(* IEC 61131-3 sources: twincat-st/tests/fixtures/negative, 10 files *)

(* ---- cp8_change_detect.st ---- *)
FUNCTION_BLOCK FB_ChangeDetect
VAR_INPUT
  fSetpoint  : LREAL;  // [mm]
  bStart    : BOOL;
END_VAR
VAR_OUTPUT
  bSetpointChanged : BOOL;
END_VAR
VAR
  fTarget    : LREAL;  // [mm] setpoint latched at start
END_VAR
IF bStart THEN
  fTarget := fSetpoint;
END_IF
bSetpointChanged := (fTarget <> fSetpoint);
END_FUNCTION_BLOCK

(* ---- FB_AbstractHook.st ---- *)
// CP24 must stay quiet on the abstract method's parameter: it has no body to use
// it in, by design. The concrete method's parameter is used and also stays quiet.
FUNCTION_BLOCK ABSTRACT FB_AbstractHook
VAR_OUTPUT
    nLast : INT;
END_VAR

METHOD ABSTRACT OnStep
VAR_INPUT
    nStep : INT;
END_VAR

METHOD Record
VAR_INPUT
    nValue : INT;
END_VAR
nLast := nValue;

(* ---- FB_ConditionalCallsClean.st ---- *)
// X12, CP7 and CP12 must stay quiet on every shape here. A timer reset with
// IN := FALSE on the way into its state, blocks called unconditionally, an Error
// bound with '=>', read as a member, or handed on whole, and an output written in
// both branches of one IF are all correct.
FUNCTION_BLOCK FB_ConditionalCallsClean
VAR_INPUT
    bStart   : BOOL;
    bSensor  : BOOL;
    fPos     : LREAL;    // mm
END_VAR
VAR_OUTPUT
    bFault   : BOOL;
END_VAR
VAR
    eStep    : E_Step;
    tonWait  : TON;
    tonStep  : TON;
    fbEdge   : R_TRIG;
    fbMove   : MC_MoveAbsolute;
    fbPower  : MC_Power;
    fbHome   : MC_Home;
    axisX    : AXIS_REF;
    bMoveErr : BOOL;
    qbValve AT %Q* : BOOL;
END_VAR
fbEdge(CLK := bSensor);
tonStep(IN := eStep = E_Step.Settle, PT := T#500MS);
CASE eStep OF
    E_Step.Idle:
        IF bStart THEN
            tonWait(IN := FALSE);   // lint:allow CP20 the reset on the way into Wait
            eStep := E_Step.Wait;
        END_IF
    E_Step.Wait:
        tonWait(IN := TRUE, PT := T#2S);
        IF tonWait.Q OR fbEdge.Q THEN
            eStep := E_Step.Settle;
        END_IF
    E_Step.Settle:
        IF tonStep.Q THEN
            eStep := E_Step.Idle;
        END_IF
    E_Step.Error:
        eStep := E_Step.Idle;
ELSE
    eStep := E_Step.Error;
END_CASE
fbPower(Axis := axisX, Enable := TRUE);
fbMove(Axis := axisX, Execute := eStep = E_Step.Settle, Position := fPos,
       Velocity := 50.0, Error => bMoveErr);
fbHome(Axis := axisX, Execute := bStart);
IF bMoveErr OR fbPower.Error THEN
    qbValve := FALSE;
ELSE
    qbValve := eStep = E_Step.Wait;
END_IF
bFault := CheckHome(fbHome);
END_FUNCTION_BLOCK

METHOD CheckHome : BOOL
VAR_IN_OUT
    fbBlock : MC_Home;
END_VAR
CheckHome := fbBlock.Error;
END_METHOD

(* ---- FB_GuardedTimer.st ---- *)
// X12 stays silent on two guards TcOpen calls its task timers in: one entered
// whenever the timer's input drops ('... OR NOT bIn'), so the call there resets it,
// and one that only checks the reference the preset is read through. CP24 stays
// silent on a variable XAE declared for a UML state chart, which only the chart uses.
FUNCTION_BLOCK FB_GuardedTimer
VAR_INPUT
    bIn         : BOOL;
    bUseTimeout : BOOL;
    tTimeout    : TIME;
END_VAR
VAR_IN_OUT
    refCfg : ST_TimerCfg;
END_VAR
VAR_OUTPUT
    bTimedOut : BOOL;
    bInfo     : BOOL;
END_VAR
VAR
    {attribute 'hide'}
    fbTimer : TON;
    {attribute 'hide'}
    fbInfo : TON;
    {attribute 'implicit_state_chart_struct' := ''}
    UML_SC_Main : _UML_SC_0123456789abcdef0123456789abcdef;
    rCfg : REFERENCE TO ST_TimerCfg;
END_VAR
rCfg REF= refCfg;
IF bUseTimeout OR NOT bIn THEN
    fbTimer(IN := bIn, PT := tTimeout);
END_IF
IF __ISVALIDREF(rCfg) THEN
    fbInfo(IN := bIn, PT := rCfg.tInfo);
END_IF
bTimedOut := fbTimer.Q;
bInfo := fbInfo.Q;
END_FUNCTION_BLOCK

(* ---- FB_RefBinding.st ---- *)
// 'REF=' binds a reference; it compares nothing, so CP8 and CP28 stay silent.
// The bound members sit behind pragma lines, as in the library that showed it.
FUNCTION_BLOCK FB_RefBinding
VAR_OUTPUT
    tActive : TIME;
    fActive : LREAL;
END_VAR
VAR
    {attribute 'hide'}
    tSlow : TIME := T#5S;
    {attribute 'hide'}
    fGain : LREAL := 1.5;
    rTime : REFERENCE TO TIME;
    rGain : REFERENCE TO LREAL;
END_VAR
rTime REF= tSlow;
rGain REF= fGain;
IF __ISVALIDREF(rTime) AND __ISVALIDREF(rGain) THEN
    tActive := rTime;
    fActive := rGain;
END_IF
END_FUNCTION_BLOCK

(* ---- FB_RefOrder.st ---- *)
// E3: an ordering comparison through a REFERENCE TO, or through a dereferenced
// pointer, is on the values behind them, not on addresses. A reference is
// dereferenced implicitly and p^ is the value, so none of these is E3. Field
// round 4 reported 'ist_Zone.fEnd <= ist_Zone.fStart' (two LREAL members read
// through a REFERENCE TO a zone struct) as high, twice, on a production project.
FUNCTION_BLOCK FB_RefOrder
VAR_INPUT
    ist_Zone : REFERENCE TO ST_Zone;    // fStart, fEnd : LREAL [mm]
    refA : REFERENCE TO LREAL;
    refB : REFERENCE TO LREAL;
    pZone : POINTER TO ST_Zone;
    pA : POINTER TO LREAL;
    pB : POINTER TO LREAL;
END_VAR
VAR_OUTPUT
    bEmpty : BOOL;
    bBelow : BOOL;
    bPtrEmpty : BOOL;
    bPtrBelow : BOOL;
END_VAR
// Members read through a reference: the shape the field reported.
IF __ISVALIDREF(ist_Zone) THEN
    bEmpty := ist_Zone.fEnd <= ist_Zone.fStart;
END_IF
// Two references compared directly: still the values.
IF __ISVALIDREF(refA) THEN
    IF __ISVALIDREF(refB) THEN
        bBelow := refA < refB;
    END_IF
END_IF
// Members and values read through a dereferenced pointer.
IF pZone <> 0 THEN
    bPtrEmpty := pZone^.fEnd <= pZone^.fStart;
END_IF
IF pA <> 0 THEN
    IF pB <> 0 THEN
        bPtrBelow := pA^ < pB^;
    END_IF
END_IF
END_FUNCTION_BLOCK

(* ---- FB_RemanentMode.st ---- *)
// X13 stays silent. A remembered operating mode is chosen by the operator, not
// stepped by its own CASE, and a remanent part counter selects nothing. The step
// counter of the sequence is a plain VAR, the shape Rule 9 asks for.
FUNCTION_BLOCK FB_RemanentMode
VAR_INPUT
    nModeRequest : INT;
    bPart        : BOOL;
    bStart       : BOOL;
END_VAR
VAR_OUTPUT
    fSpeed : LREAL;
    bError : BOOL;
END_VAR
VAR PERSISTENT
    nMode      : INT;
    nPartCount : UDINT;
END_VAR
VAR
    nStep  : INT;
    fbPart : R_TRIG;
END_VAR
IF nModeRequest > 0 THEN
    nMode := nModeRequest;
END_IF
CASE nMode OF
    1: fSpeed := 0.5;
    2: fSpeed := 1.0;
ELSE
    fSpeed := 0.0;
END_CASE
fbPart(CLK := bPart);
IF fbPart.Q THEN
    nPartCount := nPartCount + 1;
END_IF
CASE nStep OF
    0:  IF bStart THEN nStep := 10; END_IF
    10: IF NOT bStart THEN nStep := 0; END_IF
    99: bError := TRUE;
        IF NOT bStart THEN bError := FALSE; nStep := 0; END_IF
ELSE
    nStep := 99;
END_CASE
END_FUNCTION_BLOCK

(* ---- FB_SecondaryCase.st ---- *)
// X7 and X3 must stay quiet on the second CASE. It only picks a value per step,
// a step without a label keeps the last one on purpose, and the state variable it
// reads has an error state and an ELSE in the main CASE above it.
FUNCTION_BLOCK FB_SecondaryCase
VAR_INPUT
    bStart : BOOL;
    bReset : BOOL;
END_VAR
VAR_OUTPUT
    bError : BOOL;
END_VAR
VAR
    eStep   : E_Step;
    fTarget : LREAL;   // [mm]
END_VAR
CASE eStep OF
    E_Step.Idle:
        IF bStart THEN
            eStep := E_Step.Move;
        END_IF
    E_Step.Move:
        eStep := E_Step.Idle;
    E_Step.DeviceError:
        bError := TRUE;
        IF bReset THEN
            bError := FALSE;
            eStep := E_Step.Idle;
        END_IF
ELSE
    eStep := E_Step.DeviceError;
END_CASE

CASE eStep OF
    E_Step.Idle:
        fTarget := 0.0;
    E_Step.Move:
        fTarget := 120.0;
END_CASE
END_FUNCTION_BLOCK

(* ---- FB_StepExecute.st ---- *)
// X11 must stay quiet on every Execute here. A step comparison is edge-correct
// because the step changes; a trigger's .Q is an edge by construction; a lone
// command bit is set and cleared by whoever owns it, which the text cannot judge.
FUNCTION_BLOCK FB_StepExecute
VAR_INPUT
    bStart  : BOOL;
    bEnable : BOOL;
    bJog    : BOOL;
    fPos    : LREAL;
    fVelo   : LREAL;
END_VAR
VAR_OUTPUT
    bFault  : BOOL;
END_VAR
VAR
    eStep    : E_Step;
    fbMove   : MC_MoveAbsolute;
    fbJog    : MC_MoveVelocity;
    fbHome   : MC_Home;
    fbTrig   : R_TRIG;
    bHomeCmd : BOOL;
    axisX    : AXIS_REF;
END_VAR
fbTrig(CLK := bJog);
fbMove(Axis := axisX, Execute := (eStep = E_Step.Move) AND bEnable, Position := fPos,
       Velocity := fVelo);
fbJog(Axis := axisX, Execute := fbTrig.Q AND bEnable, Velocity := fVelo);
fbHome(Axis := axisX, Execute := bHomeCmd);
fbHome.Execute := bStart;
bFault := fbMove.Error OR fbJog.Error OR fbHome.Error;
END_FUNCTION_BLOCK

(* ---- x7_secondary_case.st ---- *)
TYPE E_Step :
(
  Idle    := 0,
  MoveA    := 10,
  MoveB    := 20,
  DeviceError  := 900
);
END_TYPE

FUNCTION_BLOCK FB_TwoCases
VAR_INPUT
  bGo      : BOOL;
  bFault    : BOOL;
  bReset    : BOOL;
END_VAR
VAR
  eStep    : E_Step;
  fTarget    : LREAL;  // [mm]
END_VAR
IF bFault THEN
  eStep := E_Step.DeviceError;
END_IF
CASE eStep OF
  E_Step.Idle:    IF bGo THEN eStep := E_Step.MoveA; END_IF
  E_Step.MoveA:    eStep := E_Step.MoveB;
  E_Step.MoveB:    eStep := E_Step.Idle;
  E_Step.DeviceError:  IF bReset THEN eStep := E_Step.Idle; END_IF
ELSE
  eStep := E_Step.DeviceError;
END_CASE
// Pick a target per step; other steps keep the last one
CASE eStep OF
  E_Step.MoveA:  fTarget := 100.0;
  E_Step.MoveB:  fTarget := 0.0;
END_CASE
END_FUNCTION_BLOCK
